// TIA Portal V20 export
DATA_BLOCK "02_Wartungsfreigaben_DB"   // DB22
// stored: InstanceOfName 02_Wartungsfreigaben, InstanceOfType FB
"02_Wartungsfreigaben"
   // VAR
   //    Tag_Result : Word;
   //    Status_F_PWD : Bool;
   //    Status_FULL_PWD : Bool;
   //    Status_R_PWD : Bool;
   //    Status_HMI_PWD : Bool;
   //    REQ : Bool;
   //    F_PWD : Bool;
   //    FULL_PWD : Bool;
   //    R_PWD : Bool;
   //    HMI_PWD : Bool;
   //    TP_REQ : TP_TIME;
   //    "F-Wartungsfreigabe_freigeben" : Bool;
   //    "F-Wartungsfreigabe_sperren" : Bool;
   //    "FULL-Wartungsfreigabe_freigeben" : Bool;
   //    "FULL-Wartungsfreigabe_sperren" : Bool;
   // END_VAR
BEGIN
END_DATA_BLOCK
